(* IEC 61131-3 sources: Gen-AI/release/member2-v1.1/成员2_提交包_v1.1/agent/logs/scenario_fixture/repair/fixture/E3_S01_1_42, 3 files *)

(* ---- best.st ---- *)
FUNCTION_BLOCK FB_S01
VAR_INPUT
    StartBtn : BOOL;
    LeftPartPresent : BOOL;
    RightPartPresent : BOOL;
    EStop_NC : BOOL;
END_VAR
VAR_OUTPUT
    ClampLeft : BOOL;
    ClampRight : BOOL;
    Busy : BOOL;
    Status : WORD;
END_VAR
(* Add a VAR block for internal state/timers before the implementation, if needed. *)
(* SKELETON ONLY: replace this RETURN with scan logic and required initial state. *)
RETURN;
END_FUNCTION_BLOCK

(*  *)

(* ---- final.st ---- *)
FUNCTION_BLOCK FB_S01
VAR_INPUT
    StartBtn : BOOL;
    LeftPartPresent : BOOL;
    RightPartPresent : BOOL;
    EStop_NC : BOOL;
END_VAR
VAR_OUTPUT
    ClampLeft : BOOL;
    ClampRight : BOOL;
    Busy : BOOL;
    Status : WORD;
END_VAR
(* Add a VAR block for internal state/timers before the implementation, if needed. *)
(* SKELETON ONLY: replace this RETURN with scan logic and required initial state. *)
RETURN;
END_FUNCTION_BLOCK

(*  *)

(* ---- skeleton.st ---- *)
FUNCTION_BLOCK FB_S01
VAR_INPUT
    StartBtn : BOOL;
    LeftPartPresent : BOOL;
    RightPartPresent : BOOL;
    EStop_NC : BOOL;
END_VAR
VAR_OUTPUT
    ClampLeft : BOOL;
    ClampRight : BOOL;
    Busy : BOOL;
    Status : WORD;
END_VAR
(* Add a VAR block for internal state/timers before the implementation, if needed. *)
(* SKELETON ONLY: replace this RETURN with scan logic and required initial state. *)
RETURN;
END_FUNCTION_BLOCK
